RoboDK station: Bench V1 cell v3.rdk

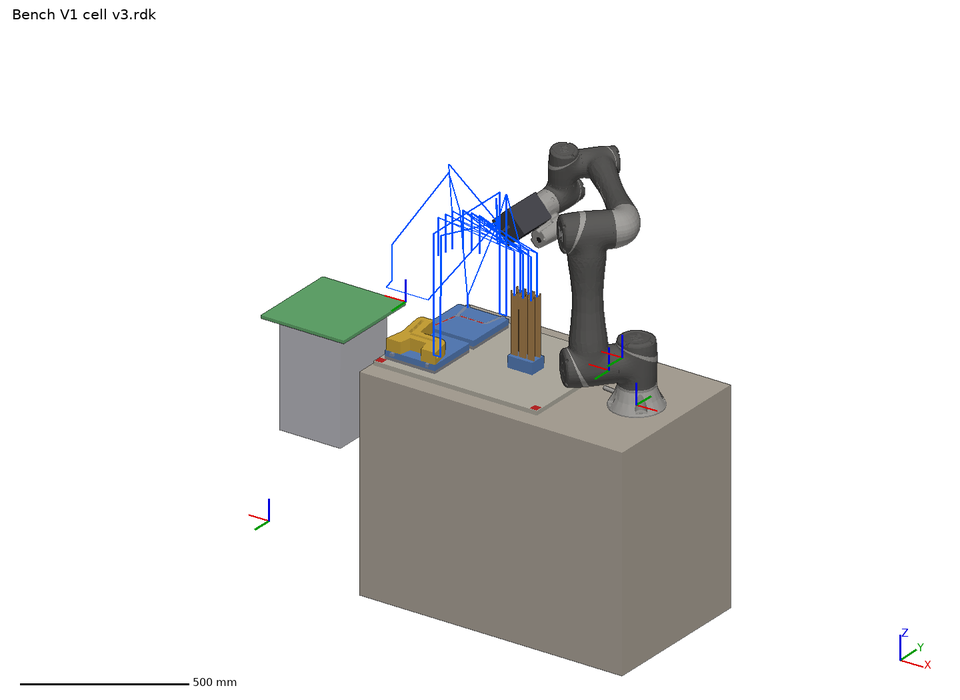
[picture v0: the station drawn from its stored meshes, robots at their saved joint values, targets as dots, program paths as lines]
Station Bench V1 cell v3 (saved by RoboDK 6.1.1). Poses are relative to the parent item; angles as X-Y-Z fixed-axis rotations.
  - frame Cell at (0, 0, 0) mm
    - frame Work plate at (-206.44, 152.99, -4.46) mm, rotated rx -0.03 ry -0.07 rz -179.98 deg
      - frame Ground base at (0, -67, 15) mm
        - object Table at (0, 0, 0) mm, size 950 x 560 x 735 mm
        - object Ground base plate at (0, 0, 0) mm, size 590 x 440 x 15 mm, geometry from ground_base.stl
        - object Vision square 1 at (3, 3, 0) mm, size 25 x 25 x 0.5 mm, geometry from vision_square.stl
        - object Vision square 2 at (562, 3, 0) mm, size 25 x 25 x 0.5 mm, geometry from vision_square.stl
        - object Vision square 3 at (3, 412, 0) mm, size 25 x 25 x 0.5 mm, geometry from vision_square.stl
        - object Vision square 4 at (562, 412, 0) mm, size 25 x 25 x 0.5 mm, geometry from vision_square.stl
        - object Base A riser at (480, 120, 10) mm, size 180 x 180 x 10 mm
        - object Base A at (480, 120, 10) mm, size 180 x 180 x 20 mm, geometry from base_a.stl
        - object Base B riser at (480, 320, 10) mm, size 180 x 180 x 10 mm
        - object Base B at (480, 320, 10) mm, size 180 x 180 x 20 mm, geometry from base_b.stl
        - object Plank jig at (150, 190, 0) mm, size 90 x 60 x 40 mm, geometry from plank_jig.stl
        - frame AMR at (740, 60, 0) mm
          - object AMR plate at (0, 0, 0) mm, size 300 x 320 x 10 mm
          - object AMR top module at (0, 0, 0) mm, size 220 x 240 x 372 mm
          - frame Omron LD-250 Base at (380, 160, -765) mm
            - robot AMR LD-250: 4 axes
                joint limits [-10000, -10000, -10, -3600] to [10000, 10000, 10, 3600]; home [0, 0, 0, 0]; saved at [0, 0, 0, 0]
        - object frame1 at (477.29, 93.12, 144.5) mm, rotated rx 0 ry 0 rz -90 deg, size 174.7 x 141.9 x 10 mm, geometry from frame.stl
        - object frame2 at (477.29, 346.88, -95.5) mm, rotated rx 180 ry 0 rz 90 deg, size 174.7 x 141.9 x 10 mm, geometry from frame.stl
        - object piece A1 at (477.29, 98.12, 144.5) mm, rotated rx 90 ry 0 rz 0 deg, size 21.4 x 10 x 5 mm, geometry from interface_piece.stl
        - object piece B1 at (477.29, 341.88, 144.5) mm, rotated rx 90 ry 0 rz -180 deg, size 21.4 x 10 x 5 mm, geometry from interface_piece.stl
        - object plank1 at (165, 207.5, 125) mm, rotated rx 90 ry 0 rz 0 deg, size 25 x 250 x 5 mm, geometry from plank_body.stl
        - object piece A2 at (447.3, 98.12, 144.5) mm, rotated rx 90 ry 0 rz 0 deg, size 21.4 x 10 x 5 mm, geometry from interface_piece.stl
        - object piece B2 at (447.3, 341.88, 144.5) mm, rotated rx 90 ry 0 rz -180 deg, size 21.4 x 10 x 5 mm, geometry from interface_piece.stl
        - object plank2 at (195, 207.5, 125) mm, rotated rx 90 ry 0 rz 0 deg, size 25 x 250 x 5 mm, geometry from plank_body.stl
        - object piece A3 at (507.27, 98.12, 144.5) mm, rotated rx 90 ry 0 rz 0 deg, size 21.4 x 10 x 5 mm, geometry from interface_piece.stl
        - object piece B3 at (507.27, 341.88, 144.5) mm, rotated rx 90 ry 0 rz -180 deg, size 21.4 x 10 x 5 mm, geometry from interface_piece.stl
        - object plank3 at (225, 207.5, 125) mm, rotated rx 90 ry 0 rz 0 deg, size 25 x 250 x 5 mm, geometry from plank_body.stl
        - object piece A4 at (529.24, 116.56, 144.5) mm, rotated rx 90 ry 0 rz 80 deg, size 21.4 x 10 x 5 mm, geometry from interface_piece.stl
        - object piece B4 at (529.24, 323.44, 144.5) mm, rotated rx 90 ry 0 rz 100 deg, size 21.4 x 10 x 5 mm, geometry from interface_piece.stl
        - object plank4 at (165, 237.5, 125) mm, rotated rx 90 ry 0 rz 0 deg, size 25 x 250 x 5 mm, geometry from plank_body.stl
        - object piece A5 at (534.45, 146.09, 144.5) mm, rotated rx 90 ry 0 rz 80 deg, size 21.4 x 10 x 5 mm, geometry from interface_piece.stl
        - object piece B5 at (534.45, 293.91, 144.5) mm, rotated rx 90 ry 0 rz 100 deg, size 21.4 x 10 x 5 mm, geometry from interface_piece.stl
        - object plank5 at (195, 237.5, 125) mm, rotated rx 90 ry 0 rz 0 deg, size 25 x 250 x 5 mm, geometry from plank_body.stl
        - object piece A6 at (539.66, 175.62, 144.5) mm, rotated rx 90 ry 0 rz 80 deg, size 21.4 x 10 x 5 mm, geometry from interface_piece.stl
        - object piece B6 at (539.66, 264.38, 144.5) mm, rotated rx 90 ry 0 rz 100 deg, size 21.4 x 10 x 5 mm, geometry from interface_piece.stl
        - object plank6 at (225, 237.5, 125) mm, rotated rx 90 ry 0 rz 0 deg, size 25 x 250 x 5 mm, geometry from plank_body.stl
        - object Guide at (480, 320, 90) mm, rotated rx 180 ry 0 rz 0 deg, size 177.7 x 180 x 40 mm, geometry from guide.stl
        - target Home (Cartesian target) at (295, 220, 380) mm, rotated rx 180 ry 0 rz 0 deg; joints [-14.089, 2.917, -80.099, -12.747, -90.01, 75.887] of Omron TM5-900
        - target guide B-A pick out low (Cartesian target) at (383, 390, 50) mm, rotated rx 0 ry 90 rz 0 deg; joints [8.389, -22.724, -132.74, -24.469, 98.365, 89.963] of Omron TM5-900
        - target guide B-A pick out (Cartesian target) at (383, 390, 450) mm, rotated rx 0 ry 90 rz 0 deg; joints [8.433, 10.061, -100.143, -89.851, 98.409, 89.963] of Omron TM5-900
        - target guide B-A via (Cartesian target) at (295, 220, 450) mm, rotated rx 0 ry 90 rz 0 deg; joints [-32.59, 30.389, -113.158, -97.152, 57.386, 90.016] of Omron TM5-900
        - target guide B-A wrist ready (Cartesian target) at (295, 220, 380) mm, rotated rx -104.58 ry -32.51 rz -35.36 deg; joints [-50.728, 20.278, -116.455, -24.612, -14.272, 24.981] of Omron TM5-900
        - target guide B-A wrist swapped (joint target) at (338.91, 166.36, 496.05) mm, rotated rx -75.5 ry -32.53 rz -66.1 deg; joints [-50.728, 20.278, -116.455, -24.612, 14.272, 24.981] of Omron TM5-900
        - target guide B-A via (Cartesian target) at (295, 220, 450) mm, rotated rx 0 ry 90 rz 0 deg; joints [-32.59, 30.389, -113.158, -97.152, 57.386, 90.016] of Omron TM5-900
        - target guide B-A pick (Cartesian target) at (408, 390, 50) mm, rotated rx 0 ry 90 rz 0 deg; joints [7.812, -24.505, -129.214, -26.214, 97.788, 89.964] of Omron TM5-900
        - target guide B-A lift (Cartesian target) at (408, 390, 70) mm, rotated rx 0 ry 90 rz 0 deg; joints [7.814, -21.463, -128.95, -29.52, 97.79, 89.964] of Omron TM5-900
        - target guide B-A up (Cartesian target) at (408, 390, 450) mm, rotated rx 0 ry 90 rz 0 deg; joints [7.851, 6.883, -97.45, -89.366, 97.827, 89.964] of Omron TM5-900
        - target guide B-A across (Cartesian target) at (408, 50, 450) mm, rotated rx 0 ry 90 rz 0 deg; joints [-45.328, 6.909, -97.45, -89.364, 44.648, 90.04] of Omron TM5-900
        - target guide B-A place (Cartesian target) at (408, 50, 50) mm, rotated rx 0 ry -90 rz -180 deg; joints [-45.297, -24.479, -129.215, -26.212, 44.679, -89.96] of Omron TM5-900
        - target guide B-A over place (Cartesian target) at (408, 50, 450) mm, rotated rx 0 ry -90 rz -180 deg; joints [-45.328, 6.909, -97.45, -89.364, 44.648, -89.96] of Omron TM5-900
        - target guide B-A place approach (Cartesian target) at (408, 50, 90) mm, rotated rx 0 ry -90 rz -180 deg; joints [-45.3, -18.508, -128.521, -32.876, 44.676, -89.96] of Omron TM5-900
        - target guide B-A place out (Cartesian target) at (383, 50, 50) mm, rotated rx 0 ry -90 rz -180 deg; joints [-48.296, -22.696, -132.741, -24.463, 41.68, -89.952] of Omron TM5-900
        - target guide B-A place out up (Cartesian target) at (383, 50, 450) mm, rotated rx 0 ry -90 rz -180 deg; joints [-48.333, 10.089, -100.144, -89.845, 41.642, -89.952] of Omron TM5-900
        - target plank3 pick travel (Cartesian target) at (225, 205, 380) mm, rotated rx 180 ry 0 rz -90 deg; joints [-18.429, 12.369, -88.214, -14.084, -90.005, -198.454] of Omron TM5-900
        - target plank3 pick approach (Cartesian target) at (225, 205, 275) mm, rotated rx 180 ry 0 rz -90 deg; joints [-18.431, 14.063, -104.285, 0.293, -90.005, -198.455] of Omron TM5-900
        - target plank3 pick (Cartesian target) at (225, 205, 235) mm, rotated rx 180 ry 0 rz -90 deg; joints [-18.431, 13.759, -109.643, 5.956, -90.005, -198.455] of Omron TM5-900
        - target plank3 pick out (Cartesian target) at (225, 205, 295) mm, rotated rx 180 ry 0 rz -90 deg; joints [-18.43, 14.01, -101.456, -2.482, -90.005, -198.454] of Omron TM5-900
        - target plank3 pick up (Cartesian target) at (225, 205, 380) mm, rotated rx 180 ry 0 rz -90 deg; joints [-18.429, 12.369, -88.214, -14.084, -90.005, -198.454] of Omron TM5-900
        - target plank3 place travel (Cartesian target) at (507.27, 95.62, 380) mm, rotated rx 180 ry 0 rz -90 deg; joints [-19.585, -31.821, -35.961, -22.146, -90.003, -199.609] of Omron TM5-900
        - target plank3 above guide (Cartesian target) at (507.27, 95.62, 329.5) mm, rotated rx 180 ry 0 rz -90 deg; joints [-19.585, -28.774, -48.091, -13.064, -90.003, -199.609] of Omron TM5-900
        - target plank3 place (Cartesian target) at (507.27, 95.62, 254.5) mm, rotated rx 180 ry 0 rz -90 deg; joints [-19.585, -27.192, -61.018, -1.719, -90.003, -199.609] of Omron TM5-900
        - target plank3 push approach (Cartesian target) at (507.27, 95.62, 289.5) mm, rotated rx 180 ry 0 rz -90 deg; joints [-19.585, -27.6, -55.517, -6.811, -90.003, -199.609] of Omron TM5-900
        - target plank3 push (Cartesian target) at (507.27, 95.62, 269.5) mm, rotated rx 180 ry 0 rz -90 deg; joints [-19.585, -27.304, -58.757, -3.867, -90.003, -199.609] of Omron TM5-900
        - target plank3 push out (Cartesian target) at (507.27, 95.62, 289.5) mm, rotated rx 180 ry 0 rz -90 deg; joints [-19.585, -27.6, -55.517, -6.811, -90.003, -199.609] of Omron TM5-900
        - target plank3 place up (Cartesian target) at (507.27, 95.62, 380) mm, rotated rx 180 ry 0 rz -90 deg; joints [-19.585, -31.821, -35.961, -22.146, -90.003, -199.609] of Omron TM5-900
        - target plank6 pick travel (Cartesian target) at (225, 235, 380) mm, rotated rx 180 ry 0 rz -90 deg; joints [-14.439, 12.367, -88.214, -14.082, -90.01, -194.463] of Omron TM5-900
        - target plank6 pick approach (Cartesian target) at (225, 235, 275) mm, rotated rx 180 ry 0 rz -90 deg; joints [-14.441, 14.061, -104.285, 0.295, -90.01, -194.465] of Omron TM5-900
        - target plank6 pick (Cartesian target) at (225, 235, 235) mm, rotated rx 180 ry 0 rz -90 deg; joints [-14.442, 13.757, -109.644, 5.958, -90.01, -194.466] of Omron TM5-900
        - target plank6 pick out (Cartesian target) at (225, 235, 295) mm, rotated rx 180 ry 0 rz -90 deg; joints [-14.441, 14.009, -101.457, -2.481, -90.01, -194.465] of Omron TM5-900
        - target plank6 pick up (Cartesian target) at (225, 235, 380) mm, rotated rx 180 ry 0 rz -90 deg; joints [-14.439, 12.367, -88.214, -14.082, -90.01, -194.463] of Omron TM5-900
        - target plank6 place travel (Cartesian target) at (542.12, 175.18, 380) mm, rotated rx 180 ry 0 rz -10 deg; joints [-12.785, -37.947, -25.826, -26.156, -90.012, 87.191] of Omron TM5-900
        - target plank6 above guide (Cartesian target) at (542.12, 175.18, 329.5) mm, rotated rx 180 ry 0 rz -10 deg; joints [-12.785, -33.547, -40.655, -15.727, -90.012, 87.191] of Omron TM5-900
        - target plank6 place (Cartesian target) at (542.12, 175.18, 254.5) mm, rotated rx 180 ry 0 rz -10 deg; joints [-12.787, -31.253, -54.883, -3.793, -90.012, 87.189] of Omron TM5-900
        - target plank6 push approach (Cartesian target) at (542.12, 175.18, 289.5) mm, rotated rx 180 ry 0 rz -10 deg; joints [-12.786, -31.919, -48.939, -9.071, -90.012, 87.19] of Omron TM5-900
        - target plank6 push (Cartesian target) at (542.12, 175.18, 269.5) mm, rotated rx 180 ry 0 rz -10 deg; joints [-12.786, -31.466, -52.456, -6.008, -90.012, 87.19] of Omron TM5-900
        - target plank6 push out (Cartesian target) at (542.12, 175.18, 289.5) mm, rotated rx 180 ry 0 rz -10 deg; joints [-12.786, -31.919, -48.939, -9.071, -90.012, 87.19] of Omron TM5-900
        - target plank6 place up (Cartesian target) at (542.12, 175.18, 380) mm, rotated rx 180 ry 0 rz -10 deg; joints [-12.785, -37.947, -25.826, -26.156, -90.012, 87.191] of Omron TM5-900
        - target plank2 pick travel (Cartesian target) at (195, 205, 380) mm, rotated rx 180 ry 0 rz -90 deg; joints [-19.849, 16.424, -91.186, -15.166, -90.003, 160.127] of Omron TM5-900
        - target plank2 pick approach (Cartesian target) at (195, 205, 275) mm, rotated rx 180 ry 0 rz -90 deg; joints [-19.85, 18.419, -107.374, -0.973, -90.003, 160.126] of Omron TM5-900
        - target plank2 pick (Cartesian target) at (195, 205, 235) mm, rotated rx 180 ry 0 rz -90 deg; joints [-19.85, 18.235, -112.832, 4.668, -90.003, 160.126] of Omron TM5-900
        - target plank2 pick out (Cartesian target) at (195, 205, 295) mm, rotated rx 180 ry 0 rz -90 deg; joints [-19.85, 18.305, -104.507, -3.726, -90.003, 160.126] of Omron TM5-900
        - target plank2 pick up (Cartesian target) at (195, 205, 380) mm, rotated rx 180 ry 0 rz -90 deg; joints [-19.849, 16.424, -91.186, -15.166, -90.003, 160.127] of Omron TM5-900
        - target plank2 place travel (Cartesian target) at (447.3, 95.62, 380) mm, rotated rx 180 ry 0 rz -90 deg; joints [-21.345, -20.954, -52.182, -16.792, -90.001, 158.631] of Omron TM5-900
        - target plank2 above guide (Cartesian target) at (447.3, 95.62, 329.5) mm, rotated rx 180 ry 0 rz -90 deg; joints [-21.345, -19.166, -61.856, -8.907, -90.001, 158.631] of Omron TM5-900
        - target plank2 place (Cartesian target) at (447.3, 95.62, 254.5) mm, rotated rx 180 ry 0 rz -90 deg; joints [-21.345, -18.495, -73.245, 1.812, -90.001, 158.631] of Omron TM5-900
        - target plank2 push approach (Cartesian target) at (447.3, 95.62, 289.5) mm, rotated rx 180 ry 0 rz -90 deg; joints [-21.345, -18.55, -68.29, -3.088, -90.001, 158.631] of Omron TM5-900
        - target plank2 push (Cartesian target) at (447.3, 95.62, 269.5) mm, rotated rx 180 ry 0 rz -90 deg; joints [-21.345, -18.467, -71.191, -0.27, -90.001, 158.631] of Omron TM5-900
        - target plank2 push out (Cartesian target) at (447.3, 95.62, 289.5) mm, rotated rx 180 ry 0 rz -90 deg; joints [-21.345, -18.55, -68.29, -3.088, -90.001, 158.631] of Omron TM5-900
        - target plank2 place up (Cartesian target) at (447.3, 95.62, 380) mm, rotated rx 180 ry 0 rz -90 deg; joints [-21.345, -20.954, -52.182, -16.792, -90.001, 158.631] of Omron TM5-900
        - target plank5 pick travel (Cartesian target) at (195, 235, 380) mm, rotated rx 180 ry 0 rz -90 deg; joints [-15.56, 16.422, -91.186, -15.164, -90.008, 164.416] of Omron TM5-900
        - target plank5 pick approach (Cartesian target) at (195, 235, 275) mm, rotated rx 180 ry 0 rz -90 deg; joints [-15.562, 18.416, -107.374, -0.971, -90.008, 164.414] of Omron TM5-900
        - target plank5 pick (Cartesian target) at (195, 235, 235) mm, rotated rx 180 ry 0 rz -90 deg; joints [-15.563, 18.233, -112.832, 4.67, -90.008, 164.413] of Omron TM5-900
        - target plank5 pick out (Cartesian target) at (195, 235, 295) mm, rotated rx 180 ry 0 rz -90 deg; joints [-15.561, 18.303, -104.507, -3.724, -90.008, 164.415] of Omron TM5-900
        - target plank5 pick up (Cartesian target) at (195, 235, 380) mm, rotated rx 180 ry 0 rz -90 deg; joints [-15.56, 16.422, -91.186, -15.164, -90.008, 164.416] of Omron TM5-900
        - target plank5 place travel (Cartesian target) at (536.91, 145.66, 380) mm, rotated rx 180 ry 0 rz -10 deg; joints [-15.108, -37.171, -27.15, -25.608, -90.009, 84.868] of Omron TM5-900
        - target plank5 above guide (Cartesian target) at (536.91, 145.66, 329.5) mm, rotated rx 180 ry 0 rz -10 deg; joints [-15.109, -32.984, -41.552, -15.393, -90.009, 84.867] of Omron TM5-900
        - target plank5 place (Cartesian target) at (536.91, 145.66, 254.5) mm, rotated rx 180 ry 0 rz -10 deg; joints [-15.11, -30.786, -55.602, -3.541, -90.009, 84.866] of Omron TM5-900
        - target plank5 push approach (Cartesian target) at (536.91, 145.66, 289.5) mm, rotated rx 180 ry 0 rz -10 deg; joints [-15.109, -31.418, -49.717, -8.794, -90.009, 84.866] of Omron TM5-900
        - target plank5 push (Cartesian target) at (536.91, 145.66, 269.5) mm, rotated rx 180 ry 0 rz -10 deg; joints [-15.11, -30.985, -53.197, -5.747, -90.009, 84.866] of Omron TM5-900
        - target plank5 push out (Cartesian target) at (536.91, 145.66, 289.5) mm, rotated rx 180 ry 0 rz -10 deg; joints [-15.109, -31.418, -49.717, -8.794, -90.009, 84.866] of Omron TM5-900
        - target plank5 place up (Cartesian target) at (536.91, 145.66, 380) mm, rotated rx 180 ry 0 rz -10 deg; joints [-15.108, -37.171, -27.15, -25.608, -90.009, 84.868] of Omron TM5-900
        - target plank1 pick travel (Cartesian target) at (165, 205, 380) mm, rotated rx 180 ry 0 rz -90 deg; joints [-21.51, 20.489, -93.86, -16.558, -90.001, 158.466] of Omron TM5-900
        - target plank1 pick approach (Cartesian target) at (165, 205, 275) mm, rotated rx 180 ry 0 rz -90 deg; joints [-21.51, 22.877, -110.195, -2.609, -90.001, 158.466] of Omron TM5-900
        - target plank1 pick (Cartesian target) at (165, 205, 235) mm, rotated rx 180 ry 0 rz -90 deg; joints [-21.51, 22.858, -115.763, 2.976, -90.001, 158.466] of Omron TM5-900
        - target plank1 pick out (Cartesian target) at (165, 205, 295) mm, rotated rx 180 ry 0 rz -90 deg; joints [-21.51, 22.681, -107.284, -5.326, -90.001, 158.466] of Omron TM5-900
        - target plank1 pick up (Cartesian target) at (165, 205, 380) mm, rotated rx 180 ry 0 rz -90 deg; joints [-21.51, 20.489, -93.86, -16.558, -90.001, 158.466] of Omron TM5-900
        - target plank1 place travel (Cartesian target) at (477.29, 95.62, 380) mm, rotated rx 180 ry 0 rz -90 deg; joints [-20.428, -26.039, -44.868, -19.022, -90.002, 159.548] of Omron TM5-900
        - target plank1 above guide (Cartesian target) at (477.29, 95.62, 329.5) mm, rotated rx 180 ry 0 rz -90 deg; joints [-20.428, -23.785, -55.44, -10.703, -90.002, 159.548] of Omron TM5-900
        - target plank1 place (Cartesian target) at (477.29, 95.62, 254.5) mm, rotated rx 180 ry 0 rz -90 deg; joints [-20.428, -22.746, -67.427, 0.244, -90.002, 159.548] of Omron TM5-900
        - target plank1 push approach (Cartesian target) at (477.29, 95.62, 289.5) mm, rotated rx 180 ry 0 rz -90 deg; joints [-20.428, -22.948, -62.259, -4.722, -90.002, 159.548] of Omron TM5-900
        - target plank1 push (Cartesian target) at (477.29, 95.62, 269.5) mm, rotated rx 180 ry 0 rz -90 deg; joints [-20.428, -22.777, -65.292, -1.859, -90.002, 159.548] of Omron TM5-900
        - target plank1 push out (Cartesian target) at (477.29, 95.62, 289.5) mm, rotated rx 180 ry 0 rz -90 deg; joints [-20.428, -22.948, -62.259, -4.722, -90.002, 159.548] of Omron TM5-900
        - target plank1 place up (Cartesian target) at (477.29, 95.62, 380) mm, rotated rx 180 ry 0 rz -90 deg; joints [-20.428, -26.039, -44.868, -19.022, -90.002, 159.548] of Omron TM5-900
        - target plank4 pick travel (Cartesian target) at (165, 235, 380) mm, rotated rx 180 ry 0 rz -90 deg; joints [-16.873, 20.487, -93.86, -16.555, -90.006, 163.103] of Omron TM5-900
        - target plank4 pick approach (Cartesian target) at (165, 235, 275) mm, rotated rx 180 ry 0 rz -90 deg; joints [-16.875, 22.874, -110.196, -2.607, -90.006, 163.101] of Omron TM5-900
        - target plank4 pick (Cartesian target) at (165, 235, 235) mm, rotated rx 180 ry 0 rz -90 deg; joints [-16.876, 22.856, -115.763, 2.979, -90.006, 163.1] of Omron TM5-900
        - target plank4 pick out (Cartesian target) at (165, 235, 295) mm, rotated rx 180 ry 0 rz -90 deg; joints [-16.875, 22.679, -107.285, -5.323, -90.006, 163.101] of Omron TM5-900
        - target plank4 pick up (Cartesian target) at (165, 235, 380) mm, rotated rx 180 ry 0 rz -90 deg; joints [-16.873, 20.487, -93.86, -16.555, -90.006, 163.103] of Omron TM5-900
        - target plank4 place travel (Cartesian target) at (531.7, 116.13, 380) mm, rotated rx 180 ry 0 rz -10 deg; joints [-17.431, -36.736, -27.886, -25.307, -90.006, 82.545] of Omron TM5-900
        - target plank4 above guide (Cartesian target) at (531.7, 116.13, 329.5) mm, rotated rx 180 ry 0 rz -10 deg; joints [-17.431, -32.661, -42.063, -15.205, -90.006, 82.545] of Omron TM5-900
        - target plank4 place (Cartesian target) at (531.7, 116.13, 254.5) mm, rotated rx 180 ry 0 rz -10 deg; joints [-17.432, -30.517, -56.013, -3.399, -90.006, 82.544] of Omron TM5-900
        - target plank4 push approach (Cartesian target) at (531.7, 116.13, 289.5) mm, rotated rx 180 ry 0 rz -10 deg; joints [-17.432, -31.13, -50.162, -8.637, -90.006, 82.544] of Omron TM5-900
        - target plank4 push (Cartesian target) at (531.7, 116.13, 269.5) mm, rotated rx 180 ry 0 rz -10 deg; joints [-17.432, -30.709, -53.62, -5.599, -90.006, 82.544] of Omron TM5-900
        - target plank4 push out (Cartesian target) at (531.7, 116.13, 289.5) mm, rotated rx 180 ry 0 rz -10 deg; joints [-17.432, -31.13, -50.162, -8.637, -90.006, 82.544] of Omron TM5-900
        - target plank4 place up (Cartesian target) at (531.7, 116.13, 380) mm, rotated rx 180 ry 0 rz -10 deg; joints [-17.431, -36.736, -27.886, -25.307, -90.006, 82.545] of Omron TM5-900
        - target guide A-B pick out low (Cartesian target) at (383, 50, 50) mm, rotated rx 0 ry -90 rz -180 deg; joints [-48.296, -22.696, -132.741, -24.463, 41.68, -89.952] of Omron TM5-900
        - target guide A-B pick out (Cartesian target) at (383, 50, 450) mm, rotated rx 0 ry -90 rz -180 deg; joints [-48.333, 10.089, -100.144, -89.845, 41.642, -89.952] of Omron TM5-900
        - target guide A-B via (Cartesian target) at (295, 220, 450) mm, rotated rx 0 ry -90 rz -180 deg; joints [-32.59, 30.389, -113.158, -97.152, 57.386, -89.984] of Omron TM5-900
        - target guide A-B wrist ready (Cartesian target) at (531.71, 116.13, 380) mm, rotated rx -104.88 ry -18.77 rz -29.9 deg; joints [-39.321, -20.298, -77.773, -9.49, -14.759, 52.436] of Omron TM5-900
        - target guide A-B wrist swapped (joint target) at (564.45, 89.34, 513.12) mm, rotated rx -75.16 ry -18.77 rz -48.78 deg; joints [-39.321, -20.298, -77.773, -9.491, 14.759, 52.436] of Omron TM5-900
        - target guide A-B via (Cartesian target) at (295, 220, 450) mm, rotated rx 0 ry -90 rz -180 deg; joints [-32.59, 30.389, -113.158, -97.152, 57.386, -89.984] of Omron TM5-900
        - target guide A-B pick (Cartesian target) at (408, 50, 50) mm, rotated rx 0 ry -90 rz -180 deg; joints [-45.297, -24.479, -129.215, -26.212, 44.679, -89.96] of Omron TM5-900
        - target guide A-B lift (Cartesian target) at (408, 50, 70) mm, rotated rx 0 ry -90 rz -180 deg; joints [-45.298, -21.437, -128.951, -29.518, 44.678, -89.96] of Omron TM5-900
        - target guide A-B up (Cartesian target) at (408, 50, 450) mm, rotated rx 0 ry -90 rz -180 deg; joints [-45.328, 6.909, -97.45, -89.364, 44.648, -89.96] of Omron TM5-900
        - target guide A-B across (Cartesian target) at (408, 390, 450) mm, rotated rx 0 ry -90 rz -180 deg; joints [7.851, 6.883, -97.45, -89.366, 97.827, -90.036] of Omron TM5-900
        - target guide A-B place (Cartesian target) at (408, 390, 50) mm, rotated rx 0 ry 90 rz 0 deg; joints [7.812, -24.505, -129.214, -26.214, 97.788, 89.964] of Omron TM5-900
        - target guide A-B over place (Cartesian target) at (408, 390, 450) mm, rotated rx 0 ry 90 rz 0 deg; joints [7.851, 6.883, -97.45, -89.366, 97.827, 89.964] of Omron TM5-900
        - target guide A-B place approach (Cartesian target) at (408, 390, 90) mm, rotated rx 0 ry 90 rz 0 deg; joints [7.816, -18.534, -128.521, -32.878, 97.792, 89.964] of Omron TM5-900
        - target guide A-B place out (Cartesian target) at (383, 390, 50) mm, rotated rx 0 ry 90 rz 0 deg; joints [8.389, -22.724, -132.74, -24.469, 98.365, 89.963] of Omron TM5-900
        - target guide A-B place out up (Cartesian target) at (383, 390, 450) mm, rotated rx 0 ry 90 rz 0 deg; joints [8.433, 10.061, -100.143, -89.851, 98.409, 89.963] of Omron TM5-900
        - target sub pick (Cartesian target) at (540.8, 23.3, 22) mm, rotated rx -120 ry 0 rz 9.93 deg; joints [-36.46, -73.895, -17.579, -49.907, -53.325, 25.436] of Omron TM5-900
        - target sub pick approach (Cartesian target) at (540.8, 23.3, 62) mm, rotated rx -120 ry 0 rz 9.93 deg; joints [-36.46, -74.48, -10.825, -56.077, -53.326, 25.435] of Omron TM5-900
        - target sub via (Cartesian target) at (295, 220, 450) mm, rotated rx -120 ry 0 rz 9.93 deg; joints [-35.279, -15.9, -56.713, -68.206, -52.406, 26.366] of Omron TM5-900
        - target sub centre (Cartesian target) at (295, 220, 450) mm, rotated rx 0 ry 90 rz 0 deg; joints [-32.59, 30.389, -113.158, -97.152, 57.386, 90.016] of Omron TM5-900
        - target sub start wrist ready (Cartesian target) at (295, 220, 450) mm, rotated rx 0 ry 90 rz 25 deg; joints [-50.744, 22.08, -108.673, -93.281, 14.232, 90.072] of Omron TM5-900
        - target sub start wrist swapped (joint target) at (209.75, 324.41, 449.85) mm, rotated rx 0 ry 90 rz 53.46 deg; joints [-50.744, 22.08, -108.673, -93.281, -14.231, 90.072] of Omron TM5-900
        - target sub to middle (joint target) at (430, 220, 450) mm, rotated rx -120 ry 0 rz 9.93 deg; joints [-28.865, -39.901, -20.638, -76.748, -47.557, 31.854] of Omron TM5-900
        - target sub wrist ready (Cartesian target) at (430, 220, 450) mm, rotated rx -98.01 ry -11.5 rz -23.96 deg; joints [-37.562, -12.266, -74.557, -59.684, -14.31, 20.984] of Omron TM5-900
        - target sub wrist swapped (joint target) at (519.65, 151.03, 524.65) mm, rotated rx -82.03 ry -11.51 rz -51.2 deg; joints [-37.562, -12.266, -74.557, -59.684, 14.31, 20.983] of Omron TM5-900
        - target sub place (Cartesian target) at (540.8, 416.7, 267) mm, rotated rx 60 ry 0 rz -9.93 deg; joints [20.85, -81.114, -28.985, 61.645, 138.058, 40.091] of Omron TM5-900
        - target sub above guide (Cartesian target) at (540.8, 416.7, 342) mm, rotated rx 60 ry 0 rz -9.93 deg; joints [20.854, -74.914, -30.845, 57.309, 138.056, 40.086] of Omron TM5-900
        - target sub flipped (Cartesian target) at (540.8, 416.7, 387) mm, rotated rx 60 ry 0 rz -9.93 deg; joints [20.856, -72.042, -30.214, 53.807, 138.054, 40.083] of Omron TM5-900
        - target sub place out (Cartesian target) at (544.53, 438.03, 254.5) mm, rotated rx 60 ry 0 rz -9.93 deg; joints [22.031, -87.305, -18.07, 57.884, 137.268, 38.788] of Omron TM5-900
        - target sub clear (Cartesian target) at (394.53, 438.03, 254.5) mm, rotated rx 60 ry 0 rz -9.93 deg; joints [26.213, -65.651, -65.413, 86.666, 134.358, 34.476] of Omron TM5-900
        - target sub back to middle (Cartesian target) at (295, 220, 450) mm, rotated rx 60 ry 0 rz -9.93 deg; joints [11.416, -24.337, -106.582, 73.148, 143.748, 52.064] of Omron TM5-900
        - target back wrist ready (Cartesian target) at (295, 220, 450) mm, rotated rx -79.86 ry -14.65 rz -42.51 deg; joints [-50.675, 5.466, -130.579, 82.327, 14.556, 123.206] of Omron TM5-900
        - target back wrist swapped (joint target) at (358.95, 141.79, 356.29) mm, rotated rx -100.21 ry -14.66 rz -58.87 deg; joints [-50.675, 5.467, -130.579, 82.327, -14.556, 123.206] of Omron TM5-900
        - target back home (Cartesian target) at (295, 220, 380) mm, rotated rx 180 ry 0 rz 0 deg; joints [-14.089, 2.917, -80.099, -12.747, -90.01, 75.887] of Omron TM5-900
    - frame Omron TM5-900 Base at (0, 0, 0) mm
      - robot Omron TM5-900: 6 axes, payload 4 kg, reach 900 mm, repeatability 0.05 mm, weight 22.6 kg
          modified DH rows (alpha deg, a mm, theta deg, d mm): 0, 0, 0, 145.2; 90, 0, 90, 0; 0, 429, 0, 0; 0, 411, -90, 122.3; -90, 0, 0, 106.5; 90, 0, 180, 114.15
          joint limits [-270, -180, -155, -180, -180, -270] to [270, 180, 155, 180, 180, 270]; home [0, 0, 90, -90, 90, 0]; saved at [-42.131, -4.294, -82.971, -82.899, -35.224, 50.65]
        - tool EGP, TCP at (0, 0, 160) mm, size 94 x 90 x 160 mm
  - program AssembleBench (255 instructions, listed below)
  - Python program Deliver (AMR) (listed below)
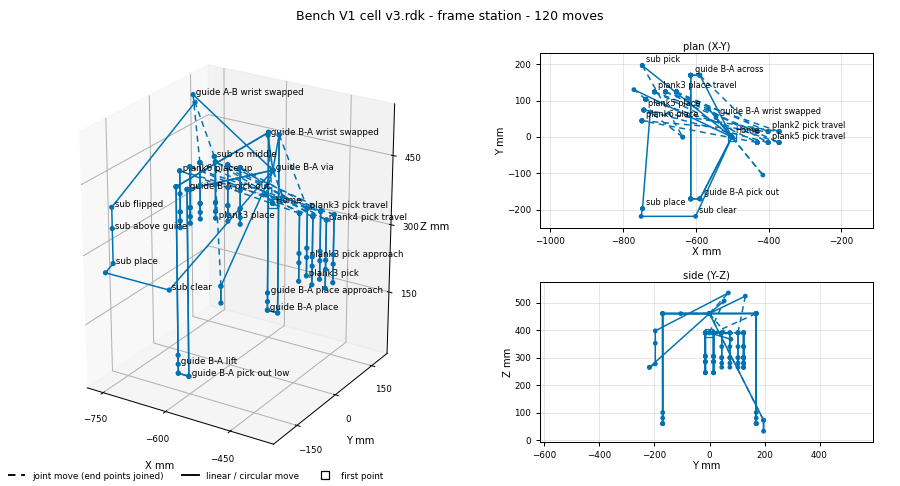
[picture p0: tool path of Bench V1 cell v3.rdk in frame station, 120 of 120 moves have a stored position in this frame; points joined in program order, loops and branches not executed]

--- program AssembleBench (robot Omron TM5-900) ---
  Simulation: parts to start
  Set Ref.: Ground base
  Set Tool: EGP
  Smooth(0)
  Set speed (100.0 mm/s)
  MoveJ (Home)
  MoveL (guide B-A wrist ready)
  MoveJ (guide B-A wrist swapped)
  MoveL (guide B-A via)
  MoveL (guide B-A pick out)
  MoveL (guide B-A pick out low)
  Set speed (20.0 mm/s)
  Set IO_0=1
  Pause 300 ms
  MoveL (guide B-A pick)
  Set IO_0=0
  Pause 500 ms
  Simulation: attach Guide
  MoveL (guide B-A lift)
  Set speed (100.0 mm/s)
  MoveL (guide B-A up)
  MoveL (guide B-A across)
  MoveJ (guide B-A over place)
  MoveL (guide B-A place approach)
  Set speed (20.0 mm/s)
  MoveL (guide B-A place)
  Set IO_0=1
  Pause 500 ms
  Simulation: release guide
  MoveL (guide B-A place out)
  Set speed (100.0 mm/s)
  MoveL (guide B-A place out up)
  MoveJ (plank3 pick travel)
  MoveL (plank3 pick approach)
  Set speed (20.0 mm/s)
  MoveL (plank3 pick)
  Set IO_0=1
  Pause 500 ms
  Simulation: attach plank3
  MoveL (plank3 pick out)
  Set speed (100.0 mm/s)
  MoveL (plank3 pick up)
  MoveJ (plank3 place travel)
  MoveL (plank3 above guide)
  Set speed (20.0 mm/s)
  MoveL (plank3 place)
  Set IO_0=0
  Pause 500 ms
  Simulation: release plank3
  MoveL (plank3 push approach)
  Set IO_0=1
  Pause 300 ms
  MoveL (plank3 push)
  MoveL (plank3 push out)
  Set IO_0=0
  Pause 300 ms
  Set speed (100.0 mm/s)
  MoveL (plank3 place up)
  MoveJ (plank6 pick travel)
  MoveL (plank6 pick approach)
  Set speed (20.0 mm/s)
  MoveL (plank6 pick)
  Set IO_0=1
  Pause 500 ms
  Simulation: attach plank6
  MoveL (plank6 pick out)
  Set speed (100.0 mm/s)
  MoveL (plank6 pick up)
  MoveJ (plank6 place travel)
  MoveL (plank6 above guide)
  Set speed (20.0 mm/s)
  MoveL (plank6 place)
  Set IO_0=0
  Pause 500 ms
  Simulation: release plank6
  MoveL (plank6 push approach)
  Set IO_0=1
  Pause 300 ms
  MoveL (plank6 push)
  MoveL (plank6 push out)
  Set IO_0=0
  Pause 300 ms
  Set speed (100.0 mm/s)
  MoveL (plank6 place up)
  MoveJ (plank2 pick travel)
  MoveL (plank2 pick approach)
  Set speed (20.0 mm/s)
  MoveL (plank2 pick)
  Set IO_0=1
  Pause 500 ms
  Simulation: attach plank2
  MoveL (plank2 pick out)
  Set speed (100.0 mm/s)
  MoveL (plank2 pick up)
  MoveJ (plank2 place travel)
  MoveL (plank2 above guide)
  Set speed (20.0 mm/s)
  MoveL (plank2 place)
  Set IO_0=0
  Pause 500 ms
  Simulation: release plank2
  MoveL (plank2 push approach)
  Set IO_0=1
  Pause 300 ms
  MoveL (plank2 push)
  MoveL (plank2 push out)
  Set IO_0=0
  Pause 300 ms
  Set speed (100.0 mm/s)
  MoveL (plank2 place up)
  MoveJ (plank5 pick travel)
  MoveL (plank5 pick approach)
  Set speed (20.0 mm/s)
  MoveL (plank5 pick)
  Set IO_0=1
  Pause 500 ms
  Simulation: attach plank5
  MoveL (plank5 pick out)
  Set speed (100.0 mm/s)
  MoveL (plank5 pick up)
  MoveJ (plank5 place travel)
  MoveL (plank5 above guide)
  Set speed (20.0 mm/s)
  MoveL (plank5 place)
  Set IO_0=0
  Pause 500 ms
  Simulation: release plank5
  MoveL (plank5 push approach)
  Set IO_0=1
  Pause 300 ms
  MoveL (plank5 push)
  MoveL (plank5 push out)
  Set IO_0=0
  Pause 300 ms
  Set speed (100.0 mm/s)
  MoveL (plank5 place up)
  MoveJ (plank1 pick travel)
  MoveL (plank1 pick approach)
  Set speed (20.0 mm/s)
  MoveL (plank1 pick)
  Set IO_0=1
  Pause 500 ms
  Simulation: attach plank1
  MoveL (plank1 pick out)
  Set speed (100.0 mm/s)
  MoveL (plank1 pick up)
  MoveJ (plank1 place travel)
  MoveL (plank1 above guide)
  Set speed (20.0 mm/s)
  MoveL (plank1 place)
  Set IO_0=0
  Pause 500 ms
  Simulation: release plank1
  MoveL (plank1 push approach)
  Set IO_0=1
  Pause 300 ms
  MoveL (plank1 push)
  MoveL (plank1 push out)
  Set IO_0=0
  Pause 300 ms
  Set speed (100.0 mm/s)
  MoveL (plank1 place up)
  MoveJ (plank4 pick travel)
  MoveL (plank4 pick approach)
  Set speed (20.0 mm/s)
  MoveL (plank4 pick)
  Set IO_0=1
  Pause 500 ms
  Simulation: attach plank4
  MoveL (plank4 pick out)
  Set speed (100.0 mm/s)
  MoveL (plank4 pick up)
  MoveJ (plank4 place travel)
  MoveL (plank4 above guide)
  Set speed (20.0 mm/s)
  MoveL (plank4 place)
  Set IO_0=0
  Pause 500 ms
  Simulation: release plank4
  MoveL (plank4 push approach)
  Set IO_0=1
  Pause 300 ms
  MoveL (plank4 push)
  MoveL (plank4 push out)
  Set IO_0=0
  Pause 300 ms
  Set speed (100.0 mm/s)
  MoveL (plank4 place up)
  MoveL (guide A-B wrist ready)
  MoveJ (guide A-B wrist swapped)
  MoveL (guide A-B via)
  MoveL (guide A-B pick out)
  MoveL (guide A-B pick out low)
  Set speed (20.0 mm/s)
  Set IO_0=1
  Pause 300 ms
  MoveL (guide A-B pick)
  Set IO_0=0
  Pause 500 ms
  Simulation: attach Guide
  MoveL (guide A-B lift)
  Set speed (100.0 mm/s)
  MoveL (guide A-B up)
  MoveL (guide A-B across)
  MoveJ (guide A-B over place)
  MoveL (guide A-B place approach)
  Set speed (20.0 mm/s)
  MoveL (guide A-B place)
  Set IO_0=1
  Pause 500 ms
  Simulation: release guide
  MoveL (guide A-B place out)
  Set speed (100.0 mm/s)
  MoveL (guide A-B place out up)
  MoveL (sub centre)
  MoveL (sub start wrist ready)
  MoveJ (sub start wrist swapped)
  MoveJ (sub via)
  MoveL (sub pick approach)
  Set speed (20.0 mm/s)
  MoveL (sub pick)
  Set IO_0=1
  Pause 500 ms
  Simulation: attach frame1
  Simulation: attach plank1
  Simulation: attach plank2
  Simulation: attach plank3
  Simulation: attach plank4
  Simulation: attach plank5
  Simulation: attach plank6
  Simulation: attach piece A1
  Simulation: attach piece A2
  Simulation: attach piece A3
  Simulation: attach piece A4
  Simulation: attach piece A5
  Simulation: attach piece A6
  MoveL (sub pick approach)
  Set speed (100.0 mm/s)
  MoveJ (sub to middle)
  MoveL (sub wrist ready)
  MoveJ (sub wrist swapped)
  MoveL (sub flipped)
  MoveL (sub above guide)
  Set speed (20.0 mm/s)
  MoveL (sub place)
  Set IO_0=0
  Pause 500 ms
  Simulation: release frame 1 with the planks
  MoveL (sub place out)
  MoveL (sub clear)
  MoveL (sub back to middle)
  Set speed (100.0 mm/s)
  MoveL (back wrist ready)
  MoveJ (back wrist swapped)
  MoveL (back home)

--- Python program Deliver (AMR) ---
"""The AMR drives the finished bench 2 m away along the table and comes back (RoboDK station script
"Deliver (AMR)").

    python robot_cell/amr_drive.py           also works from outside RoboDK

Needs only the robodk package. Everything under the station's "AMR" frame rides along: its plate,
top module and LD-250, and the bench once the robot program has set it down there (the program's
release puts the bench under the AMR frame).
"""
import time

from robodk import robolink, robomath

DISTANCE = 2000          # mm, along the ground base's x (away from the robot)
STEPS = 120              # per direction
PAUSE = 1.0              # s at the far end
OWN = ("AMR plate", "AMR top module")


def main():
    RDK = robolink.Robolink()
    amr = RDK.Item("AMR", robolink.ITEM_TYPE_FRAME)
    if not amr.Valid():
        raise SystemExit("no AMR in the open station")
    riding = [c for c in amr.Childs() if c.Type() == robolink.ITEM_TYPE_OBJECT and c.Name() not in OWN]
    home = amr.Pose()
    for out in (True, False):
        for i in range(1, STEPS + 1):
            s = i / STEPS if out else 1 - i / STEPS
            s = 0.5 - 0.5 * robomath.cos(robomath.pi * s)        # smooth start and stop
            amr.setPose(robomath.transl(DISTANCE * s, 0, 0) * home)
            RDK.Render(True)
            time.sleep(0.02)
        if out:
            time.sleep(PAUSE)
    amr.setPose(home)
    print(f"AMR drove {DISTANCE / 1000:.0f} m and back with {len(riding)} parts on its plate")


if __name__ == "__main__":
    main()
